// #24 step 3a: stage of FB_MonetTelescopeControl._ParkTelescope (property ParkStage). The values are the stage numbers of
// 0.12.0 and earlier, so the log ('Parking progress: %s') and ADS watch values read as before.
{attribute 'qualified_only'}
{attribute 'strict'}
TYPE E_ParkStage :
(
	prepare := 0,			// move flags dropped; drive to the park position (untrack) or park in place (secure, #86/#87)
	untrack := 10,			// tracking of the three axes switched off
	start_move := 20,		// park targets written, MoveAxis until all three axes are busy
	wait_moves := 40,		// MoveAxis dropped per axis when its move is done, until nothing slews
	disable_axes := 60,		// axes disabled at standstill
	secure := 80,			// brake closed: covers closed, hydraulics off; waits for the covers closed
	parked := 100			// bIsParked, bPark dropped (one call), then prepare
);
END_TYPE

(* stored: Version 1.1.0.1, ProductVersion 3.1.4024.15
   DUT E_ParkStage: Id {324b041c-0e61-470d-a5ad-136002d664d6} *)
